FUNCTION_BLOCK FB_Workshop
VAR_INPUT
    bButton : BOOL;
    bSetValid : BOOL;
    bTargetOn : BOOL;
END_VAR

VAR_OUTPUT
    bLightRelay : BOOL;
END_VAR

VAR
    fbLight : FB_Light;
    bArmed : BOOL;
    bToggle : BOOL;
END_VAR

bToggle := FALSE;

IF NOT bButton THEN
    bArmed := TRUE;
ELSIF bArmed THEN
    bArmed := FALSE;
    bToggle := TRUE;
END_IF

fbLight(
    bToggle := bToggle,
    bSetValid := bSetValid,
    bTargetOn := bTargetOn
);
bLightRelay := fbLight.bOn;

END_FUNCTION_BLOCK

(* stored: Version 1.1.0.1
   POU FB_Workshop: Id {4cb4c94a-a979-4da1-85e5-4bfab4a678c9}, SpecialFunc None *)
